Fanuc KAREL source: KX00003.KL

PROGRAM KX00003
%NOLOCKGROUP
VAR
  I: INTEGER
  J: INTEGER
  B: BOOLEAN
  F: FILE
  S: STRING[80]
  P: XYZWPR
BEGIN
  OPEN FILE F ('RW', 'MD:KFSAMPLE.DT')
  WRITE F ('SAMPLE', CR)
  CLOSE FILE F
END KX00003
